// TIA Portal V21 export
// export: Created 2026-11-22T02:34:35.6339814Z, ExportSetting WithDefaults, DisplayName Totally Integrated Automation Portal, DisplayVersion V21 Update 3, DisplayName STEP 7 Professional, DisplayVersion V21 Update 3, DisplayName STEP 7 Safety, DisplayVersion V21, DisplayName Tech WebApplication, DisplayVersion V21, DisplayName WinCC Basic/Comfort/Advanced, DisplayVersion V21 Update 3, DisplayName WinCC Unified, DisplayVersion V21 Update 3
TextList "TL_Bit"  ListRange=Bit
  TextListEntry   EntryType=SingleValue, Text="Off (0)"
  TextListEntry   EntryType=SingleValue, From=1, To=1, Text="On (1)"
